# EPICS substitutions: b-55B2VNC/src/main/c++/nds3-sdn/src/main/epics/ndssdnApp/Db/DeviceTesting.substitutions
file "nds-testing.template" {
	pattern
	{	BOARDTYPE,
		BOARDTYPEIDX,
		CBS1,
		CBS2
	}
	{
		"Test",
		"0",
		"TEST",
		"TEST",
	}
}
